Fanuc KAREL source: KA00209.KL

PROGRAM KA00209
%NOLOCKGROUP
VAR
  SRC: ARRAY[4] OF XYZWPR
  DST: ARRAY[4] OF REAL
BEGIN
  DST = SRC
END KA00209
